Staubli VAL3: copy.pgx

public program copy(string x_sSource, string& x_sTarget, bool& x_bToSave)
  local num l_j
  local num l_i
begin
  trajTemp:tTrajItem[x_sTarget].nFrameIndex=trajTemp:tTrajItem[x_sSource].nFrameIndex
  trajTemp:tTrajItem[x_sTarget].nToolIndex=trajTemp:tTrajItem[x_sSource].nToolIndex
  trajTemp:tTrajItem[x_sTarget].nMoveID=trajTemp:tTrajItem[x_sSource].nMoveID
  trajTemp:tTrajItem[x_sTarget].sID=trajTemp:tTrajItem[x_sTarget].sID
  resize(trajTemp:tTrajItem[x_sTarget].pPointItem,1,size(trajTemp:tTrajItem[x_sSource].pPointItem))
  for l_i = 0 to size(trajTemp:tTrajItem[x_sSource].pPointItem)-1
    trajTemp:tTrajItem[x_sTarget].pPointItem[l_i].pParaItem.mMdesc=trajTemp:tTrajItem[x_sSource].pPointItem[l_i].pParaItem.mMdesc
    trajTemp:tTrajItem[x_sTarget].pPointItem[l_i].pParaItem.nMoveType=trajTemp:tTrajItem[x_sSource].pPointItem[l_i].pParaItem.nMoveType
    trajTemp:tTrajItem[x_sTarget].pPointItem[l_i].pPointRx=trajTemp:tTrajItem[x_sSource].pPointItem[l_i].pPointRx
    //2025.03.18 add mlc  2025.10.16 modify by liu zhengang
    trajTemp:tTrajItem[x_sTarget].pPointItem[l_i].pInter=trajTemp:tTrajItem[x_sSource].pPointItem[l_i].pInter
    trajTemp:tTrajItem[x_sTarget].pPointItem[l_i].jJointRx=trajTemp:tTrajItem[x_sSource].pPointItem[l_i].jJointRx
    for l_j = 0 to 0
      trajTemp:tTrajItem[x_sTarget].pPointItem[l_i].pParaItem.nActionIndex[l_j]=trajTemp:tTrajItem[x_sSource].pPointItem[l_i].pParaItem.nActionIndex[l_j]
      trajTemp:tTrajItem[x_sTarget].pPointItem[l_i].pParaItem.nPercentage[l_j]=trajTemp:tTrajItem[x_sSource].pPointItem[l_i].pParaItem.nPercentage[l_j]
      trajTemp:tTrajItem[x_sTarget].pPointItem[l_i].pParaItem.iIfItem.bANDOR[l_j]=(trajTemp:tTrajItem[x_sSource].pPointItem[l_i].pParaItem.iIfItem.bANDOR[l_j]==true)
    endFor
    for l_j = 0 to 2
      trajTemp:tTrajItem[x_sTarget].pPointItem[l_i].pParaItem.iIfItem.nSigType[l_j]=trajTemp:tTrajItem[x_sSource].pPointItem[l_i].pParaItem.iIfItem.nSigType[l_j]
      trajTemp:tTrajItem[x_sTarget].pPointItem[l_i].pParaItem.iIfItem.nSigIndex[l_j]=trajTemp:tTrajItem[x_sSource].pPointItem[l_i].pParaItem.iIfItem.nSigIndex[l_j]
      trajTemp:tTrajItem[x_sTarget].pPointItem[l_i].pParaItem.iIfItem.nValue[l_j]=trajTemp:tTrajItem[x_sSource].pPointItem[l_i].pParaItem.iIfItem.nValue[l_j]
    endFor
    //
    trajTemp:tTrajItem[x_sTarget].pPointItem[l_i].pParaItem.nDelay=trajTemp:tTrajItem[x_sSource].pPointItem[l_i].pParaItem.nDelay
    trajTemp:tTrajItem[x_sTarget].pPointItem[l_i].pParaItem.nSigValue=trajTemp:tTrajItem[x_sSource].pPointItem[l_i].pParaItem.nSigValue
  endFor
  x_bToSave=true
end
